(* IEC 61131-3 sources: trust-platform/examples/OSCAT/packaging_reject_pulse/non-oop/src, 3 files *)

(* ---- Configuration.st ---- *)
CONFIGURATION PackagingRejectPulseClassicConfiguration
RESOURCE Cpu0 ON PLC
    TASK MainTask (INTERVAL := T#50ms, PRIORITY := 1);
    PROGRAM Main WITH MainTask : Main;
END_RESOURCE
END_CONFIGURATION

(* ---- Main.st ---- *)
PROGRAM Main
VAR
    RejectPulse : GEN_PULSE;
    DefectDetected : BOOL := FALSE;
    RejectSolenoid : BOOL;
END_VAR

RejectPulse(ENQ := DefectDetected, PTH := T#150ms, PTL := T#500ms);
RejectSolenoid := RejectPulse.Q;
END_PROGRAM

(* ---- Tests.st ---- *)
TEST_PROGRAM PackagingRejectPulseClassicStaysLowWithoutDefect
VAR
    RejectPulse : GEN_PULSE;
END_VAR

RejectPulse(ENQ := FALSE, PTH := T#150ms, PTL := T#500ms);

ASSERT_FALSE(IN := RejectPulse.Q);
END_TEST_PROGRAM
